// TIA Portal V21 export
// export: Created 2026-11-10T19:16:30.3669997Z, ExportSetting WithDefaults, DisplayName Totally Integrated Automation Portal, DisplayVersion V21 Update 3, DisplayName STEP 7 Professional, DisplayVersion V21 Update 3, DisplayName STEP 7 Safety, DisplayVersion V21, DisplayName Tech WebApplication, DisplayVersion V21, DisplayName WinCC Basic/Comfort/Advanced, DisplayVersion V21 Update 3, DisplayName WinCC Unified, DisplayVersion V21 Update 3
DATA_BLOCK "FB_12_DB"   // DB3
VERSION : 0.1
// stored: AutoNumber true, DBAccessibleFromOPCUA true, InstanceOfName FB_12, InstanceOfType FB
"FB_12"
   // VAR_INPUT
   //    en1 : Bool;
   //    par : "UDT_12";
   // END_VAR
   // VAR_OUTPUT
   //    q : Int;
   // END_VAR
   // VAR
   //    cnt : Int;
   //    tmr { S7_SetPoint := 'True'} : TON_TIME;
   //    edge { S7_SetPoint := 'True'} : R_TRIG;
   // END_VAR
BEGIN
END_DATA_BLOCK
